(* IEC 61131-3 sources: SortJet_MasterSPS_Aufbau.fbsproj/05_Sicherheitstechnik, 4 files *)

(* ---- Durchgang_FB_V01_00_00.fb.st ---- *)
(* METADATA
{
	"v3Meta": {
		"objectGuid": "fc23c363-cc05-42cf-86d7-bbdeb020e062"
	}
}
*)
FUNCTION_BLOCK Durchgang_FB_V01_00_00
VAR_INPUT

  // BOOL
  bpFreigabeZumOeffnenDurchgang    : BOOL;
  bpDurchgangGeschlossen           : BOOL;
  bpSKGeschlossen                  : BOOL;
  bpAbschrankung_Geschlossen       : BOOL;     //Signal aus der Safety, das die Abschrankung geschlossen ist

  // WORD
  wSicherheitskreis                : WORD;

  //Baustein
  BeweglicheAbschrankung          : ZylinderPneumatik_FB_V01_00_00;

  // POINTER
  ppParameterBaustein          : REFERENCE TO Parameter_Durchgang;

END_VAR
VAR_OUTPUT

  // BOOL
  bpAnforderungZumDurchgangOffnenGestellt : BOOL;
  bpStatusDurchgangNichtGeschlossen       : BOOL;

END_VAR
VAR
  // BOOL
  blErsterZyklus     : BOOL := TRUE;

  // TRIGGER
  rtlTuerGeschlossen : R_TRIG;

  // TIMER
  tonlNotEinlass     : TON;

END_VAR
VAR

  // HARDWARE EINGÄNGE
  in_bTasterAnforderungOeffnen_1          AT %I* : BOOL;
  in_bTasterAnforderungOeffnen_2          AT %I* : BOOL;
  in_bTasterQuittierungSchliessen_1       AT %I* : BOOL;
  in_bTasterQuittierungSchliessen_2       AT %I* : BOOL;

  // HARDWARE AUSGÄNGE
  out_bLeuchteTasterAnforderungDurchgang1  AT %Q* : BOOL;
  out_bLeuchteTasterAnforderungDurchgang2  AT %Q* : BOOL;
  out_bLeuchteTasterQuittierungDurchgang1  AT %Q* : BOOL;
  out_bLeuchteTasterQuittierungDurchgang2  AT %Q* : BOOL;
  out_bDurchgangSperren                    AT %Q* : BOOL;
  out_bVerriegelungOeffnen                 AT %Q* : BOOL;
  out_bVerriegelungSchliessen              AT %Q* : BOOL;

END_VAR
//-------------------------------------------------------------------------------------------------
// Initialisierung
//-------------------------------------------------------------------------------------------------
IF ( blErsterZyklus  ) THEN
  blErsterZyklus := FALSE;

  IF bpDurchgangGeschlossen THEN
    out_bDurchgangSperren := TRUE;
    bpAnforderungZumDurchgangOffnenGestellt := FALSE;
  END_IF
END_IF

bpAbschrankung_Geschlossen:= BeweglicheAbschrankung.in_bStatusZylinderAusgefahren; // Ausgefahren = geschlossen

//-------------------------------------------------------------------------------------------------
// BAUSTEIN: EINSTELLUNGEN
//-------------------------------------------------------------------------------------------------
// Timer
tonlNotEinlass(IN := in_bTasterAnforderungOeffnen_1 OR in_bTasterAnforderungOeffnen_2, PT := T#7S);

//-------------------------------------------------------------------------------------------------
// BAUSTEIN: VERWALTUNG DER TÜREN
//-------------------------------------------------------------------------------------------------
//Anforderung zum betreten des Sicherheitskreises durch die entsprechende Tür
IF( in_bTasterAnforderungOeffnen_1 OR in_bTasterAnforderungOeffnen_2 ) THEN
  bpAnforderungZumDurchgangOffnenGestellt := TRUE;
END_IF

(* Hinweis:
   - Zuruecksetzen der Anforderung:
     => Wenn die Tuer geoeffnet wurde
     => Quittieren der Tuer
*)
IF ( in_bTasterQuittierungSchliessen_1 or in_bTasterQuittierungSchliessen_2 ) THEN
  bpAnforderungZumDurchgangOffnenGestellt := FALSE;
END_IF

// Ansteuerung der Taster-Leuchte
out_bLeuchteTasterAnforderungDurchgang1 := out_bLeuchteTasterAnforderungDurchgang2 := (( bpAnforderungZumDurchgangOffnenGestellt AND gbFlashbit05sec )
                                                                                        OR NOT out_bDurchgangSperren );

// Bewegliche Abschrankung schließen
IF ( bpFreigabeZumOeffnenDurchgang
     AND bpAnforderungZumDurchgangOffnenGestellt
     AND ppParameterBaustein.bBeweglicheAbschrankung
     AND NOT( BeweglicheAbschrankung.epStatusZylinder = eZylinderAusgefahren) )
THEN
  BeweglicheAbschrankung.bpStartAusfahren := TRUE; //Ausfahren = schließen
  BeweglicheAbschrankung.bpStartEinfahren := FALSE;//Einfahren = öffnen
ELSE
  BeweglicheAbschrankung.bpStartAusfahren := FALSE;//Ausfahren = schließen
END_IF

IF BeweglicheAbschrankung.bpDone AND BeweglicheAbschrankung.bpStartAusfahren THEN
  BeweglicheAbschrankung.bpStartAusfahren := FALSE;//Ausfahren = schließen
END_IF

// Tür oeffnen
IF ( bpFreigabeZumOeffnenDurchgang
     AND bpAnforderungZumDurchgangOffnenGestellt
     AND( bpAbschrankung_Geschlossen OR NOT (ppParameterBaustein.bBeweglicheAbschrankung) ) ) OR tonlNotEinlass.Q
THEN
  out_bDurchgangSperren := FALSE;
ELSE
  out_bDurchgangSperren := TRUE;
END_IF

// Tür wieder schließen und zurücksetzen
rtlTuerGeschlossen(CLK := ( in_bTasterQuittierungSchliessen_1 OR in_bTasterQuittierungSchliessen_2 ) AND bpDurchgangGeschlossen );
IF ( rtlTuerGeschlossen.Q  ) THEN
  bpAnforderungZumDurchgangOffnenGestellt := FALSE;
END_IF

//IF ppParameterBaustein.bBeweglicheAbschrankung AND bpDurchgangGeschlossenVerriegelt AND NOT bpAnforderungZumDurchgangOffnenGestellt THEN
IF ppParameterBaustein.bBeweglicheAbschrankung AND bpDurchgangGeschlossen
   AND NOT bpAnforderungZumDurchgangOffnenGestellt AND NOT ( BeweglicheAbschrankung.epStatusZylinder =eZylinderEingefahren) THEN
  BeweglicheAbschrankung.bpStartAusfahren := FALSE;//Ausfahren = schließen
  BeweglicheAbschrankung.bpStartEinfahren := TRUE; //Einfahren = öffnen
END_IF

IF BeweglicheAbschrankung.bpDone AND BeweglicheAbschrankung.bpStartEinfahren THEN
  BeweglicheAbschrankung.bpStartEinfahren := FALSE;//Einfahren = öffnen
END_IF

// Bolzen ausfahren lassen
IF in_bTasterQuittierungSchliessen_1 OR in_bTasterQuittierungSchliessen_2 THEN
  out_bVerriegelungSchliessen := TRUE;
  out_bVerriegelungOeffnen    := FALSE;

ELSE
  out_bVerriegelungSchliessen := out_bDurchgangSperren;
  out_bVerriegelungOeffnen    := NOT out_bDurchgangSperren;
END_IF

//-------------------------------------------------------------------------------------------------
// BAUSTEIN: AUSGAENGE
//-------------------------------------------------------------------------------------------------
// Meldung ob die Tuer geschlossen und verschlossen ist
bpStatusDurchgangNichtGeschlossen       := NOT bpSKGeschlossen;
out_bLeuchteTasterQuittierungDurchgang1 := out_bLeuchteTasterQuittierungDurchgang2 := NOT bpDurchgangGeschlossen;

// Aufruf der Unterbausteine
BeweglicheAbschrankung(bpAktivieren:=ppParameterBaustein.bBeweglicheAbschrankung, bpFreigabe := TRUE, bpReset := Job_Stationen.abpReset[apgMKSicherheiskreis[ppParameterBaustein.eZuBlockierenderSK].eaAutomatikkreis[1]]);

// Meldungen für den Unterbaustein
WatchIoControl(T#10S, ppParameterBaustein.wMeldungsNummer + 0, (BeweglicheAbschrankung.wpFehlerNr = cMELDUNG_ZYLINDER_NICHT_AUSGEFAHREN)); //Fehler beim Schließen des Durchgangs (Ausfahren)
WatchIoControl(T#10S, ppParameterBaustein.wMeldungsNummer + 1, (BeweglicheAbschrankung.wpFehlerNr = cMELDUNG_ZYLINDER_NICHT_EINGEFAHREN)); //Fehler beim Öffnen des Durchgangs (Einfahren)
END_FUNCTION_BLOCK

(* ---- Sicherheitskreis_FB.fb.st ---- *)
(* METADATA
{
	"v3Meta": {
		"objectGuid": "054ec8d1-7d35-45dd-8fed-1d9f4cdd4ae8"
	}
}
*)
FUNCTION_BLOCK Sicherheitskreis_FB
VAR_INPUT

  // BOOLEAN
  bpFreigabeStationen                   : BOOL;
  bpAnforderungSicherheitkreisAusloesen : BOOL;
  bpSicherheitskreisGeschlossenSafety   : BOOL;

END_VAR
VAR_OUTPUT

  // BOOL
  bpAnforderungSKGestellt                    : BOOL;
  bpStationenBlocken                         : BOOL;
  bpSicherheitskreisGeschlossen              : BOOL; // Hinweis: [Zeitverzoegert 2 Sekunden] Variable gibt an ob der Sicherheitskreisgeschlossen ist
  bpFreigabeZumBetretenDesSicherheitskreises : BOOL;
  bpFreigabeSafetyAusloesen                  : BOOL;
  bpFreigabeTuerenOeffnen                    : BOOL;

  // TIMER
  tonlSKFreigabe                             : TON;

END_VAR
VAR

  // TRIGGER
  rtlSKGeschlossen        : R_TRIG;
  ftlAnforderung          : F_TRIG;

  // TIMER
  tonlStationenFreigabeSK : TON;
  tonlSKGeschlossen       : TON;

END_VAR
//-------------------------------------------------------------------------------------------------
// BAUSTEIN: TIMER
//-------------------------------------------------------------------------------------------------
(* Hinweis:
   - Ueberwachung das der Sicherheitskreis wirklich geschlossen meldet
*)
tonlSKGeschlossen(IN := bpSicherheitskreisGeschlossenSafety AND NOT bpFreigabeZumBetretenDesSicherheitskreises, PT := T#2S);
tonlSKFreigabe(IN := bpFreigabeZumBetretenDesSicherheitskreises, PT := T#2S);

bpFreigabeTuerenOeffnen   := NOT bpSicherheitskreisGeschlossenSafety;//AND bpFreigabeZumBetretenDesSicherheitskreises;
bpFreigabeSafetyAusloesen := tonlSKFreigabe.Q;

//-------------------------------------------------------------------------------------------------
// BAUSTEIN: STEUERUNG SICHERHEITSKREIS
//-------------------------------------------------------------------------------------------------

(* Hinweis:
   - Anforderung zum betreten des SK
*)
bpAnforderungSKGestellt := bpAnforderungSicherheitkreisAusloesen;

tonlStationenFreigabeSK( IN:= (bpAnforderungSKGestellt AND bpFreigabeStationen ),
                         PT := t#1s);

IF ( tonlStationenFreigabeSK.Q ) THEN
  bpFreigabeZumBetretenDesSicherheitskreises := TRUE;
END_IF

ftlAnforderung( CLK := bpAnforderungSKGestellt );
IF ftlAnforderung.Q THEN
  IF bpFreigabeZumBetretenDesSicherheitskreises THEN
    bpFreigabeZumBetretenDesSicherheitskreises := FALSE;
  END_IF
END_IF

(* Hinweis:
   - Sicherheitskreis wieder schließen und zurücksetzen
*)
rtlSKGeschlossen(CLK := bpSicherheitskreisGeschlossenSafety );

IF ( rtlSKGeschlossen.Q ) THEN
  bpAnforderungSKGestellt := FALSE;
  bpFreigabeZumBetretenDesSicherheitskreises := FALSE;
END_IF

// *************************************************************************************************
// BAUSTEIN: AUSGAENGE
// *************************** **********************************************************************
(* Hinweis:
   - Ausgaenge
*)
bpStationenBlocken                  := ( bpAnforderungSKGestellt OR NOT bpSicherheitskreisGeschlossen );
bpSicherheitskreisGeschlossen       := tonlSKGeschlossen.Q; // Die Stationen dürfen erst aktiv werden, wenn alle Regler durchgeschaltet haben
END_FUNCTION_BLOCK

(* ---- Tuerschalter_FB.fb.st ---- *)
(* METADATA
{
	"v3Meta": {
		"objectGuid": "4948c423-2ad3-469d-bcc1-6cb5d4807f3f"
	}
}
*)
FUNCTION_BLOCK Tuerschalter_FB
VAR_INPUT

  // BOOL
  bpFreigabeZumOeffnenDerTuer     : BOOL;
  bpTuerRelaisQuittiert           : BOOL;
  bpWeitereTuerenGeoeffnet        : BOOL;
  bpTuerGeschlossen               : BOOL;
  in_bTasterNothaltNichtBetaetigt : BOOL := TRUE; // Oeffner - kommt von SLC (EV_ToPLC_Tueren_Nothalt_aktiv)

  // WORD
  wSicherheitskreis           : WORD;
  wMeldungsnummer             : WORD;

END_VAR
VAR_OUTPUT

  // BOOL
  bpAnforderungZumTuerOffnenGestellt : BOOL;
  bpStatusTuerNichtGeschlossen       : BOOL;
  out_bTuerZuhaltungDeaktivieren     : BOOL;

END_VAR
VAR

  // TRIGGER
  rtlTuerGeschlossen : R_TRIG;
  ftlTuerGeoeffnet   : F_TRIG;

  // TIMER
  tonlNotEinlass     : TON;

END_VAR
VAR

  // HARDWARE EINGAENGE
  in_bTasterAnforderungTuerOeffnen             : BOOL;
  in_bTasterQuittierungTuerGeschlossen         : BOOL;

  // HARDWARE AUSGAENGE
  out_bLeuchteFreigabeTuerOeffnen              : BOOL;
  out_bLeuchteTuerNichtGeschlossen             : BOOL;
  out_bLeuchteTuerNothaltAktiv                 : BOOL;

END_VAR
(* Hinweis:
   - Dieser Baustein ist für Türschalter des Herstellers Euchner
     Anmerkung:
   - Sollte Nothalt ausgeloest werden, muss die Tür mittels Not-Entriegelung [Mechanisch] geoeffnet werden
*)
//-------------------------------------------------------------------------------------------------
// BAUSTEIN: EINSTELLUNGEN
//-------------------------------------------------------------------------------------------------
// Timer
tonlNotEinlass(IN := in_bTasterAnforderungTuerOeffnen, PT := T#7S);

//-------------------------------------------------------------------------------------------------
// BAUSTEIN: VERWALTUNG DER TÜREN
//-------------------------------------------------------------------------------------------------
//Anforderung zum betreten des Sicherheitskreises durch die entsprechende Tür
IF( in_bTasterAnforderungTuerOeffnen ) THEN
  bpAnforderungZumTuerOffnenGestellt := TRUE;
END_IF

(* Hinweis:
   - Zuruecksetzen der Anforderung:
     => Wenn die Tuer geoeffnet wurde
     => Quittieren der Tuer
*)
IF ( in_bTasterQuittierungTuerGeschlossen ) THEN
  bpAnforderungZumTuerOffnenGestellt := FALSE;
END_IF

// Tür freigeben wenn sie geoeffnet wurde, obwohl sie nicht angefordert wurde

ftlTuerGeoeffnet( CLK := bgEtherCatOK AND bpTuerGeschlossen );

IF ( ftlTuerGeoeffnet.Q AND NOT in_bTasterQuittierungTuerGeschlossen ) THEN
  out_bTuerZuhaltungDeaktivieren := TRUE;
  bpAnforderungZumTuerOffnenGestellt := TRUE;
END_IF

// Ansteuerung der Taster-Leuchte
out_bLeuchteFreigabeTuerOeffnen := (( bpAnforderungZumTuerOffnenGestellt AND gbFlashbit05sec )
                                     OR out_bTuerZuhaltungDeaktivieren );

// Tür oeffnen
IF ( bpFreigabeZumOeffnenDerTuer
     AND bpAnforderungZumTuerOffnenGestellt ) OR tonlNotEinlass.Q
THEN
  out_bTuerZuhaltungDeaktivieren := TRUE;
END_IF

// Tür wieder schließen und zurücksetzen
rtlTuerGeschlossen(CLK := in_bTasterQuittierungTuerGeschlossen AND bpTuerGeschlossen );

IF ( rtlTuerGeschlossen.Q  ) THEN
  out_bTuerZuhaltungDeaktivieren := FALSE;
  bpAnforderungZumTuerOffnenGestellt := FALSE;
END_IF

//-------------------------------------------------------------------------------------------------
// BAUSTEIN: AUSGAENGE
//-------------------------------------------------------------------------------------------------
// Meldung ob die Tuer geschlossen und verschlossen ist
bpStatusTuerNichtGeschlossen     := NOT bpTuerGeschlossen OR NOT bpTuerRelaisQuittiert;

out_bLeuchteTuerNichtGeschlossen := NOT bpTuerRelaisQuittiert OR ( bpWeitereTuerenGeoeffnet AND gbFlashbit1sec );

out_bLeuchteTuerNothaltAktiv := NOT Nothalt.bpNotHaltOK;

// Meldungen
WatchIo( NOT in_bTasterNothaltNichtBetaetigt ,wMeldungsnummer );
END_FUNCTION_BLOCK

(* ---- SteuerungSicherheitskreise.prg.st ---- *)
(* METADATA
{
	"v3Meta": {
		"objectGuid": "0713858d-73c1-43e2-8e34-fbe80fbf8cab"
	}
}
*)
PROGRAM SteuerungSicherheitskreise
VAR_INPUT
  in_bTasterSKFaecherwagenQuittieren        AT %I* : BOOL; // Taster an OP fuer FW SK quittieren
  out_bLeuchtmelderSKFaecherwagenQuittieren AT %Q* : BOOL;

  bpFreigabePuffer101Ausfahren                     : BOOL;

END_VAR
VAR_OUTPUT
END_VAR
VAR

  // BOOLEAN
  ablSicherheitskreisFreigabeStation : ARRAY [cERSTE_STATION..cLETZTE_STATION] OF BOOL;
  ablSicherheitskreisFreigabeShuttle : ARRAY [cERSTES_SHUTTLE..cLETZTES_SHUTTLE] OF BOOL;
  ablSicherheitskreisFreigabeTransferShuttle : ARRAY [cERSTES_TRANSFERSHUTTLE..cLETZTES_TRANSFERSHUTTLE] OF BOOL;
  ablSicherheitskreisAnfordernExtern : ARRAY [cERSTER_SICHERHEITSKREIS..cLETZTER_SICHERHEITSKREIS] OF BOOL;

  bpPuffer101ObenAusfahren           : BOOL;
  bpPuffer103ObenAusfahren           : BOOL;
  bpPuffer102UntenAusfahren          : BOOL;
  bpPuffer104UntenAusfahren          : BOOL;
  bpPuffer101ObenEinfahren           : BOOL;
  bpPuffer103ObenEinfahren           : BOOL;
  bpPuffer102UntenEinfahren          : BOOL;
  bpPuffer104UntenEinfahren          : BOOL;

  // STEPS
  steplPuffer101ObenAusfahren        : STEPS_TE;
  steplPuffer101ObenEinfahren        : STEPS_TE;
  steplPuffer102UntenAusfahren       : STEPS_TE;
  steplPuffer102UntenEinfahren       : STEPS_TE;
  steplPuffer103ObenAusfahren        : STEPS_TE;
  steplPuffer103ObenEinfahren        : STEPS_TE;
  steplPuffer104UntenAusfahren       : STEPS_TE;
  steplPuffer104UntenEinfahren       : STEPS_TE;

  // TIMER
  tonlPuffer101ObenAusfahren         : TON;
  tonlPuffer101ObenEinfahren         : TON;
  tonlPuffer102UntenAusfahren        : TON;
  tonlPuffer102UntenEinfahren        : TON;
  tonlPuffer103ObenAusfahren         : TON;
  tonlPuffer103ObenEinfahren         : TON;
  tonlPuffer104UntenAusfahren        : TON;
  tonlPuffer104UntenEinfahren        : TON;

  // WORD
  wlIndex                            : WORD;
  wlIndexSK                          : WORD;
  wlIndexTuer                        : WORD;
  wlIndexDurchgang                   : WORD;
  wlMeldungsnummer                   : WORD;

  wlStatusPuffer101Oben_OLD          : WORD;
  wlStatusPuffer102Unten_OLD         : WORD;
  wlStatusPuffer103Oben_OLD          : WORD;
  wlStatusPuffer104Unten_OLD         : WORD;
  wlStatusTorOben_OLD                : WORD;
  wlStatusTorUnten_OLD               : WORD;

  out_bPuffer_101_Ausfahren   AT %Q* : BOOL;
  out_bPuffer_101_Einfahren   AT %Q* : BOOL;
  out_bPuffer_102_Ausfahren   AT %Q* : BOOL;
  out_bPuffer_102_Einfahren   AT %Q* : BOOL;
  out_bPuffer_103_Ausfahren   AT %Q* : BOOL;
  out_bPuffer_103_Einfahren   AT %Q* : BOOL;
  out_bPuffer_104_Ausfahren   AT %Q* : BOOL;
  out_bPuffer_104_Einfahren   AT %Q* : BOOL;

END_VAR
//-------------------------------------------------------------------------------------------------
// Aufrufe
//-------------------------------------------------------------------------------------------------
Freigabe_Stationen();
Meldungen();
Tueren();
Zuweisung_Freigabe();

// Aufruf Türen
FOR wlIndex := cERSTE_TUER TO cLETZTE_TUER DO
  aTuer[wlIndex](wMeldungsnummer := (ioccNotausAnTuer1Betaetigt - 1) + wlIndex  );
END_FOR

// Aufruf Durchgang
FOR wlIndex := cERSTER_DURCHGANG TO cLETZTER_DURCHGANG DO
  aDurchgang[wlIndex](ppParameterBaustein := (apgMKDurchgang[wlIndex]));
END_FOR

// Aufruf Sicherheitskreise
FOR wlIndex := cERSTER_SICHERHEITSKREIS TO cLETZTER_SICHERHEITSKREIS DO
  Sicherheitskreis[wlIndex]();
END_FOR
END_PROGRAM
